FUNCTION_BLOCK Pusher_IMC (* Composite Function Block Type *)
  (* Standard: 61499-2 *)
  (* Version 0.0, 10/22/2026, macie, Schneider Electric, template *)
  PACKAGE Main;
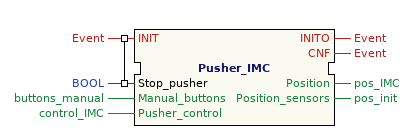
  EVENT_INPUT
    INIT WITH Stop_pusher; (* Initialization Request *)
  END_EVENT
  EVENT_OUTPUT
    INITO; (* Initialization Confirm *)
    CNF; (* Execution Confirmation *)
  END_EVENT
  VAR_INPUT
    Stop_pusher : BOOL; (* Input event qualifier *)
  END_VAR
  SOCKETS
    Manual_buttons : buttons_manual;
    Pusher_control : control_IMC;
  END_SOCKETS
  PLUGS
    Position : pos_IMC;
    Position_sensors : pos_init;
  END_PLUGS
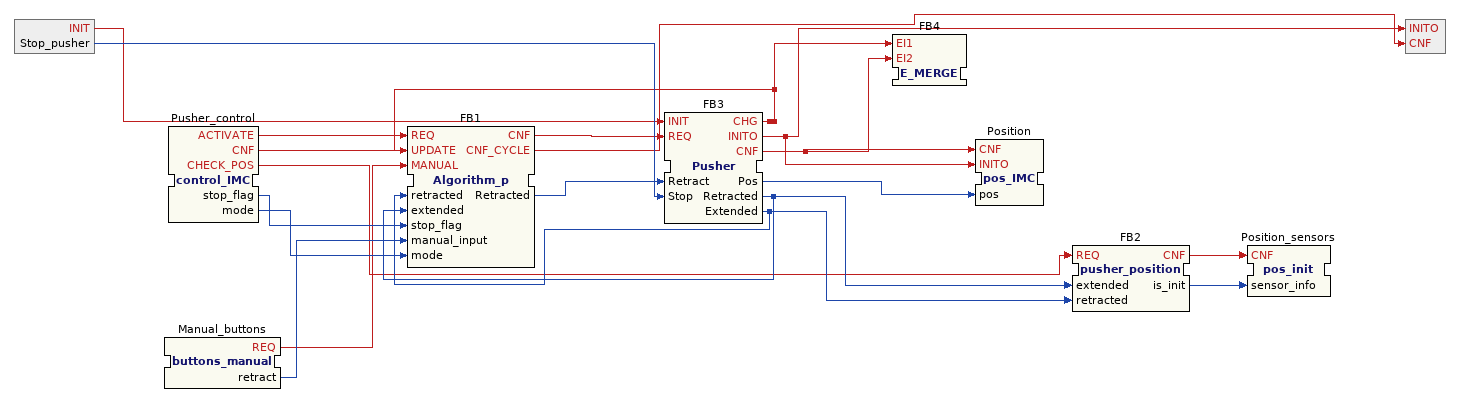
  FBS
    FB3 : Pusher;
    FB4 : E_MERGE;
    FB2 : pusher_position;
    FB1 : Algorithm_p;
  END_FBS
  EVENT_CONNECTIONS
    FB3.CHG TO FB4.EI1;
    FB3.CNF TO FB4.EI2;
    INIT TO FB3.INIT;
    FB3.INITO TO INITO;
    FB3.CNF TO Position.CNF;
    FB2.CNF TO Position_sensors.CNF;
    FB1.CNF TO FB3.REQ;
    FB3.INITO TO Position.INITO;
    FB3.CHG TO FB1.UPDATE;
    Pusher_control.ACTIVATE TO FB1.REQ;
    Pusher_control.CNF TO FB1.UPDATE;
    Manual_buttons.REQ TO FB1.MANUAL;
    FB1.CNF_CYCLE TO CNF;
    Pusher_control.CHECK_POS TO FB2.REQ;
  END_CONNECTIONS
  DATA_CONNECTIONS
    Stop_pusher TO FB3.Stop;
    FB3.Retracted TO FB2.extended;
    FB3.Extended TO FB2.retracted;
    FB3.Pos TO Position.pos;
    FB1.Retracted TO FB3.Retract;
    FB3.Retracted TO FB1.extended;
    FB3.Extended TO FB1.retracted;
    Pusher_control.stop_flag TO FB1.stop_flag;
    Pusher_control.mode TO FB1.mode;
    Manual_buttons.retract TO FB1.manual_input;
    FB2.is_init TO Position_sensors.sensor_info;
  END_CONNECTIONS
END_FUNCTION_BLOCK
